ADAPTER IWaypoint (* Adapter Interface *)
  (* Standard: 61499-1 *)
  (* Version 0.0, 11/16/2026, Sandeep Patil, Flexbridge AB *)
  PACKAGE Flexbridge.FestoMPS400;
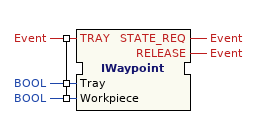
  EVENT_INPUT
    TRAY WITH Tray, Workpiece; (* To the plug: tray state changed (or answer to STATE_REQ) *)
  END_EVENT
  EVENT_OUTPUT
    STATE_REQ; (* From the plug: tell me the tray state *)
    RELEASE; (* From the plug: release the tray *)
  END_EVENT
  VAR_INPUT
    Tray : BOOL; (* A tray is at the stopper *)
    Workpiece : BOOL; (* The tray carries a workpiece *)
  END_VAR
  SERVICE SOCKET/PLUG
    SEQUENCE tray
      PLUG.STATE_REQ() -> SOCKET.STATE_REQ();
      SOCKET.TRAY(Tray, Workpiece) -> PLUG.TRAY(Tray, Workpiece);
      PLUG.RELEASE() -> SOCKET.RELEASE();
    END_SEQUENCE
  END_SERVICE
END_ADAPTER
